(* IEC 61131-3 sources: plc_simulator/plc, 4 files *)

(* ---- types.st ---- *)
USING Siemens.Simatic.Communication.OUC;
USING Siemens.Simatic.Communication.OpenUser;
USING Siemens.Simatic.Communication.MQTT;
USING Siemens.Simatic.Communication.Util;
USING System.Strings;
USING System.Serialization;

/*
#### IO map

1. control box
button: start, stop,reset
led, auto,stop,warn
errormsg

2. belt
motor command: enable, speed
motor state: state, speed

3. sensor
IR
Banner

#### Controller Main Logic
1. running state transition
idle -> running -> suspend -> stop
running -> error -> reset -> running

2. belt layout configuration
graph
link table

2. sequence start

*/

TYPE

    Station_1_Input : STRUCT
        button_1_1_1 : BOOL;
        button_1_1_2 : BOOL;
        button_1_1_3 : BOOL;
        sensor_1_1_1 : BOOL;
        button_1_2_1 : BOOL;
        button_1_2_2 : BOOL;
        button_1_2_3 : BOOL;
        sensor_1_2_1 : DWORD;
        button_1_3_1 : BOOL;
        button_1_3_2 : BOOL;
        button_1_3_3 : BOOL;
        sensor_1_3_1 : DWORD;
        clock : LINT;

    END_STRUCT;
END_TYPE

TYPE
    Station_1_Output : STRUCT
        led_1_1_1 : BOOL;
        led_1_1_2 : BOOL;
        led_1_1_3 : BOOL;
        led_1_2_1 : BOOL;
        led_1_2_2 : BOOL;
        led_1_2_3 : BOOL;
        led_1_3_1 : BOOL;
        led_1_3_2 : BOOL;
        led_1_3_3 : BOOL;

        belt_1_1_1: ARRAY[0..1] of REAL;
        belt_1_1_2: ARRAY[0..1] of REAL;
        belt_1_1_3: ARRAY[0..1] of REAL;
        belt_1_1_4: ARRAY[0..1] of REAL;
        belt_1_1_5: ARRAY[0..1] of REAL;
        // belt_1_1_6: ARRAY[0..1] of REAL;

        belt_1_2_1: ARRAY[0..1] of REAL;
        belt_1_2_2: ARRAY[0..1] of REAL;
        belt_1_2_3: ARRAY[0..1] of REAL;
        belt_1_2_4: ARRAY[0..1] of REAL;
        belt_1_2_5: ARRAY[0..1] of REAL;

        belt_1_3_1: ARRAY[0..1] of REAL;
        belt_1_3_2: ARRAY[0..1] of REAL;
        belt_1_3_3: ARRAY[0..1] of REAL;
        belt_1_3_4: ARRAY[0..1] of REAL;
        belt_1_3_5: ARRAY[0..1] of REAL;

    END_STRUCT;
END_TYPE

(* ---- tcp_client_lib.st ---- *)
USING Siemens.Simatic.Communication.OUC;
USING System;
USING System.Serialization; // For handling byte-to-integer conversions

FUNCTION TcpBlockMove
    VAR_IN_OUT
        source : ARRAY[*] OF BYTE;
        dest : ARRAY[*] OF BYTE;
    END_VAR
    VAR_INPUT
        srcOffset : UDINT;
        dstOffset : UDINT;
        count : UDINT;
    END_VAR
    VAR_TEMP
        I : UDINT;
        srcIdx : DINT;
        dstIdx : DINT;
    END_VAR

    IF count = UDINT#0 THEN
        RETURN;
    END_IF;

    srcIdx := LOWER_BOUND(source, 1) + TO_DINT(srcOffset);
    dstIdx := LOWER_BOUND(dest, 1) + TO_DINT(dstOffset);

    FOR I := UDINT#0 TO count - UDINT#1 DO
        dest[dstIdx] := source[srcIdx];
        srcIdx := srcIdx + DINT#1;
        dstIdx := dstIdx + DINT#1;
    END_FOR;
END_FUNCTION

CLASS TcpClient
    VAR CONSTANT
        MAX_SEND_LENGTH : UINT := UINT#256;
        MAX_RECEIVE_LENGTH : UINT := UINT#256;
    END_VAR

    VAR PUBLIC
        IsConfigured : BOOL := FALSE;
        IsConnected : BOOL := FALSE;

        ConnectDone, ConnectError, ConnectBusy : BOOL;
        ConnectExecute : BOOL;
        ConnectStatus, LastConnectStatus : WORD;
        ConnectAttemptCount, ConnectDoneCount, ConnectErrorCount : UDINT;

        SendDone, SendError, SendBusy : BOOL;
        SendExecute : BOOL;
        SendStatus, LastSendStatus : WORD;
        SendDoneCount, SendErrorCount, DroppedSendCount : UDINT;

        ReceiveNewData, ReceiveError, ReceiveBusy : BOOL;
        ReceiveStatus, LastReceiveStatus : WORD;
        ReceiveLength :INT;
        ReceiveCount, ReceiveErrorCount : UDINT;
        ReceiveBuffer : ARRAY [0..MAX_RECEIVE_LENGTH - UINT#1] OF BYTE;
    END_VAR

    VAR PRIVATE
        config : ConnectionConfiguration;
        connect : Connect;
        send : TcpSend;
        receive : TcpReceive;
        sendTimer : IEC.TON;
        sendPeriod : TIME := T#1S;
        sendBuffer : ARRAY [0..MAX_SEND_LENGTH - UINT#1] OF BYTE;
        sendLength : UDINT := UDINT#0;
        sendQueued : BOOL := FALSE;
        prevConnectExecute : BOOL := FALSE;
           retryTimer : IEC.TON;
    retryDelay : TIME := T#2S;
    forceExecuteLow : BOOL := FALSE;

    END_VAR

    METHOD PUBLIC Configure
        VAR_INPUT
            remoteAddress : Siemens.Simatic.Communication.IPConfiguration.IPv4;
            remotePort : UINT;
            connectionID : WORD := WORD#1;
            hardwareID : UINT := UINT#64;
            period : TIME := T#1S;
        END_VAR

        IF NOT IsConfigured THEN
            config.HardwareID := hardwareID;
            config.ConnectionID := connectionID;
            config.RemoteAddress := remoteAddress;
            config.RemotePort := remotePort;
            sendPeriod := period;
            IsConfigured := TRUE;
        END_IF;
    END_METHOD

    METHOD PUBLIC QueueSend
        VAR_INPUT
            dataLength : UDINT;
        END_VAR
        VAR_IN_OUT
            data : ARRAY[*] OF BYTE;
        END_VAR

        IF (dataLength + UDINT#8) > TO_UDINT(MAX_SEND_LENGTH) THEN
            DroppedSendCount := DroppedSendCount + UDINT#1;
            RETURN;
        END_IF;

        IF SendBusy THEN
            DroppedSendCount := DroppedSendCount + UDINT#1;
            RETURN;
        END_IF;

        sendLength := dataLength + UDINT#8;

        // Fixed magic marker 16#12345678, followed by little-endian UDINT payload length.
        sendBuffer[0] := BYTE#16#12;
        sendBuffer[1] := BYTE#16#34;
        sendBuffer[2] := BYTE#16#56;
        sendBuffer[3] := BYTE#16#78;
        sendBuffer[4] := TO_BYTE(TO_DWORD(dataLength) AND DWORD#16#FF);
        sendBuffer[5] := TO_BYTE(SHR(TO_DWORD(dataLength), USINT#8) AND DWORD#16#FF);
        sendBuffer[6] := TO_BYTE(SHR(TO_DWORD(dataLength), USINT#16) AND DWORD#16#FF);
        sendBuffer[7] := TO_BYTE(SHR(TO_DWORD(dataLength), USINT#24) AND DWORD#16#FF);

        TcpBlockMove(
            source := data,
            dest := sendBuffer,
            srcOffset := UDINT#0,
            dstOffset := UDINT#8,
            count := dataLength
        );

        sendQueued := TRUE;
    END_METHOD

    METHOD PUBLIC Run

        VAR_TEMP
            recv_len : udint;
            END_VAR

// in Run():
IF ConnectError THEN
    forceExecuteLow := TRUE;
    retryTimer(IN := TRUE, PT := retryDelay);
ELSIF retryTimer.Q THEN
    forceExecuteLow := FALSE;
    retryTimer(IN := FALSE);
END_IF;

ConnectExecute := NOT IsConnected AND NOT connect.busy AND NOT forceExecuteLow;

        IF NOT IsConfigured THEN
            RETURN;
        END_IF;

        // ConnectExecute := NOT IsConnected AND NOT connect.busy;
        IF ConnectExecute AND NOT prevConnectExecute THEN
            ConnectAttemptCount := ConnectAttemptCount + UDINT#1;
        END_IF;
        prevConnectExecute := ConnectExecute;

        // connect(
        // execute := NOT IsConnected AND NOT connect.busy,
        // connectionID := config.ConnectionID,
        // connectionConfiguration := config,
        // done => ConnectDone,
        //     busy => ConnectBusy,
        //     error => ConnectError,
        //     status => ConnectStatus
        // );

        connect(
            execute := ConnectExecute,
            connectionID := config.ConnectionID,
            connectionConfiguration := config,
            done => ConnectDone,
            busy => ConnectBusy,
            error => ConnectError,
            status => ConnectStatus
        );

        IF ConnectStatus <> WORD#16#7000 THEN
            LastConnectStatus := ConnectStatus;
        END_IF;

        IF ConnectDone THEN
            ConnectDoneCount := ConnectDoneCount + UDINT#1;
            IsConnected := TRUE;
        END_IF;

        IF ConnectError THEN
            ConnectErrorCount := ConnectErrorCount + UDINT#1;
        END_IF;

        sendTimer(IN := IsConnected AND sendQueued AND NOT sendTimer.Q, PT := sendPeriod);
        SendExecute := IsConnected AND sendQueued AND sendTimer.Q AND NOT send.busy;

        send(
            execute := SendExecute,
            connectionID := config.ConnectionID,
            length := sendLength,
            data := sendBuffer,
            done => SendDone,
            busy => SendBusy,
            error => SendError,
            status => SendStatus
        );

        IF SendStatus <> WORD#16#7000 THEN
            LastSendStatus := SendStatus;
        END_IF;

        IF SendDone THEN
            SendDoneCount := SendDoneCount + UDINT#1;
        END_IF;

        IF SendError THEN
            SendErrorCount := SendErrorCount + UDINT#1;
        END_IF;
        receive(
            enable := IsConnected,
            connectionID := config.ConnectionID,
            adhocMode := TRUE,
            data := ReceiveBuffer,
            length := MAX_RECEIVE_LENGTH,

            newDataReceived => ReceiveNewData,
            receivedLength =>  recv_len,
            busy => ReceiveBusy,
            error => ReceiveError,
            status => ReceiveStatus
        );

        IF ReceiveNewData THEN
            ReceiveLength := TO_INT(recv_len);
        ELSE
            ReceiveLength := INT#0;
        END_IF;

        IF ReceiveStatus <> WORD#16#7000 THEN
            LastReceiveStatus := ReceiveStatus;
        END_IF;

        IF ReceiveNewData THEN
            ReceiveCount := ReceiveCount + UDINT#1;
        END_IF;

        IF ReceiveError THEN
            ReceiveErrorCount := ReceiveErrorCount + UDINT#1;
        END_IF;
    END_METHOD
END_CLASS

CLASS TCP_StreamParser1

    VAR CONSTANT
        BUFFER_LENGTH : INT := 4095;
        PAYLOAD_LENGTH : INT := 2048;

        // Instance of your TRCV or communication interface
        // e.g., MyTrcvInstance : TRCV;
    END_VAR

    VAR
        // Adjust buffer size depending on your largest expected payload + 8 byte header
        Buffer : Array[0..BUFFER_LENGTH] Of Byte;
        BufferLength : Int := 0; // Tracks current number of valid bytes in Buffer

    END_VAR

    VAR PUBLIC
        // Parsing variables
        // i : Int := 0;
        MagicFound : Bool := False;
        MarkerIndex : Int := 0;
        PayloadLength : DInt := 0;
        TotalPacketSize : Int := 0;

        // Output/Export extracted data
        PayloadReady : Bool := False;
        ExtractedPayload : Array[0..PAYLOAD_LENGTH] Of Byte;
        ExtractedLength : Int := 0;
    END_VAR

    METHOD PUBLIC Execute
        VAR
            MoveIndex : Int;

        END_VAR
        VAR_IN_OUT
           // Temp array to capture immediate cycle data from network
            RxTemp : Array[*] Of Byte;
            RxCount : Int;
        END_VAR
        VAR_TEMP
            i : int;

        END_VAR

        PayloadReady := False; // Reset flag every cycle

        // 1. SIMULATED/ACTUAL RECV CALL: Fetch raw data from network interface
        // Replace this block with your actual TRCV logic
        // TRCV_Instance(RCV:=RxTemp, ...NDR=>DataReady, LEN=>RxCount);

        // If data arrived this cycle, append it to our main stream buffer
        IF RxCount > 0 THEN
            // Ensure we don't overflow our main stream buffer
            IF (BufferLength + RxCount) <= 4096 THEN
                // Copy temporary network chunk to the end of our stream buffer
                FOR i := 0 TO RxCount - 1 DO
                    Buffer[BufferLength + i] := RxTemp[i];
                END_FOR;
                BufferLength := BufferLength + RxCount;
            ELSE
                // Handle Buffer Overflow Error here (e.g., reset buffer)
                BufferLength := 0;
            END_IF;
        END_IF;

        // 2. PARSING LOOP: Process buffer continuously until no complete packets remain
        WHILE BufferLength >= 8 DO // Must have at least 8 bytes (4B Magic + 4B Length)

            MagicFound := False;

            // Look for the 4-byte Magic Marker: 0x12345678
            FOR i := 0 TO (BufferLength - 4) DO
                IF Buffer[i] = TO_BYTE(16#12) AND Buffer[i+1] = TO_BYTE(16#34) AND Buffer[i+2] = TO_BYTE(16#56) AND Buffer[i+3] = TO_BYTE(16#78) THEN
                    MagicFound := True;
                    MarkerIndex := i;
                    EXIT; // Found the earliest marker, break FOR loop
                END_IF;
            END_FOR;

            // If magic marker is not anywhere in the buffer, discard junk data safely
            IF NOT MagicFound THEN
                // Keep only the last 3 bytes in case the magic word was split between frames
                IF BufferLength > 3 THEN
                    FOR i := 0 TO 2 DO
                        Buffer[i] := Buffer[BufferLength - 3 + i];
                    END_FOR;
                    BufferLength := 3;
                END_IF;
                EXIT; // Break the WHILE loop, wait for more data
            END_IF;

            // If the magic marker was found deeper in the stream, slide buffer to align to it
            IF MarkerIndex > 0 THEN
                FOR i := 0 TO (BufferLength - 1 - MarkerIndex) DO
                    Buffer[i] := Buffer[MarkerIndex + i];
                END_FOR;
                BufferLength := BufferLength - MarkerIndex;
            END_IF;

            // Double check if we still have the full 8 bytes header after realignment
            IF BufferLength < 8 THEN
                EXIT; // Wait for next cycle data
            END_IF;

            // 3. EXTRACT LENGTH: Deserialize 4 bytes following the magic marker (little-endian)
            // Reconstructs DInt from Buffer[4..7]
            // PayloadLength := TO_DINT(SHL(TO_DWORD(Buffer[4]), UINT#24) OR
            //                  SHL(TO_DWORD(Buffer[5]), UINT#16) OR
            //                  SHL(TO_DWORD(Buffer[6]), UINT#8)  OR
            //                  TO_DWORD(Buffer[7]));

            // Combined safely into a DINT
PayloadLength := TO_DINT(
    TO_DWORD(Buffer[4]) OR
    SHL(TO_DWORD(Buffer[5]), USINT#8) OR
    SHL(TO_DWORD(Buffer[6]), USINT#16) OR
    SHL(TO_DWORD(Buffer[7]), USINT#24)
);

            TotalPacketSize := 8 + TO_INT(PayloadLength);

            // 4. CHECK COMPLETENESS: Ensure the complete payload length has arrived
            IF BufferLength < TotalPacketSize THEN
                EXIT; // Packet incomplete. Stop parsing and wait for the rest of the stream
            END_IF;

            // 5. EXTRACT PAYLOAD: Complete packet found! Copy it to output array
            FOR i := 0 TO TO_INT(PayloadLength) - 1 DO
                ExtractedPayload[i] := Buffer[8 + i];
            END_FOR;

            ExtractedLength := TO_INT(PayloadLength);
            PayloadReady := True; // Signal to consumer logic that data is ready

            // Execute application-specific logic with ExtractedPayload here if needed...

            // 6. SLIDE STREAM BUFFER: Shift remaining trailing data to index 0
            BufferLength := BufferLength - TotalPacketSize;
            IF BufferLength > 0 THEN
                FOR i := 0 TO (BufferLength - 1) DO
                    Buffer[i] := Buffer[TotalPacketSize + i];
                END_FOR;
            END_IF;

        END_WHILE;
    END_METHOD
END_CLASS

CLASS TCP_StreamParser

    VAR CONSTANT
        BUFFER_LENGTH : INT := 4095;
        PAYLOAD_LENGTH : INT := 2048;
        HEADER_SIZE : INT := 8;
    END_VAR

    VAR
        // Persistent internal stream buffer
        Buffer : Array[0..BUFFER_LENGTH] Of Byte;
        BufferLength : Int := 0; // Tracks current number of valid bytes in Buffer
    END_VAR

    VAR PUBLIC
        // Parsing state variables
        MagicFound : Bool := False;
        MarkerIndex : Int := 0;
        PayloadLength : DInt := 0;
        TotalPacketSize : Int := 0;

        // Output / Export data interface
        PayloadReady : Bool := False;
        PayloadReadyCount : Int := 0;

        ExtractedPayload : Array[0..PAYLOAD_LENGTH] Of Byte;
        ExtractedLength : Int := 0;
    END_VAR

    METHOD PUBLIC Execute
        VAR_IN_OUT
            // Dynamic bounds array to safely read variable network chunk sizes
            RxTemp : Array[*] Of Byte;
            RxCount : Int;
        END_VAR

        VAR_TEMP
            i : INT;
            UpperIndexBound : DINT;
        END_VAR

        PayloadReady := False; // Reset flag every cycle

        // 1. APPEND NEW NETWORK DATA TO STREAM BUFFER
        IF RxCount > 0 THEN
            // FIX 1: Dynamically match against the upper bound of the constant size (4095 index = 4096 size)
            IF (BufferLength + RxCount) <= (BUFFER_LENGTH + 1) THEN
                FOR i := 0 TO RxCount - 1 DO
                    Buffer[BufferLength + i] := RxTemp[LOWER_BOUND(RxTemp, 1) + TO_DINT(i)];
                END_FOR;
                BufferLength := BufferLength + RxCount;
            ELSE
                // Buffer Overflow Safety: Wipe pointer to avoid crashing the PLC PLC
                BufferLength := 0;
            END_IF;
        END_IF;

        // 2. PARSING LOOP: Process internal stream buffer
        WHILE BufferLength >= HEADER_SIZE DO

            MagicFound := False;

            // Look for the 4-byte Magic Marker: 0x12345678
            FOR i := 0 TO (BufferLength - 4) DO
                IF Buffer[i] = TO_BYTE(16#12) AND Buffer[i+1] = TO_BYTE(16#34) AND Buffer[i+2] = TO_BYTE(16#56) AND Buffer[i+3] = TO_BYTE(16#78) THEN
                    MagicFound := True;
                    MarkerIndex := i;
                    EXIT; // Found the earliest marker, break FOR loop
                END_IF;
            END_FOR;

            // FIX 2: Handle garbage data or unmatched fragments safely without losing potential split markers
            IF NOT MagicFound THEN
                IF BufferLength > 3 THEN
                    FOR i := 0 TO 2 DO
                        Buffer[i] := Buffer[BufferLength - 3 + i];
                    END_FOR;
                    BufferLength := 3;
                END_IF;
                EXIT; // Force break of WHILE loop to wait for more data
            END_IF;

            // If the magic marker was found deeper in the stream, slide buffer to align to it
            IF MarkerIndex > 0 THEN
                FOR i := 0 TO (BufferLength - 1 - MarkerIndex) DO
                    Buffer[i] := Buffer[MarkerIndex + i];
                END_FOR;
                BufferLength := BufferLength - MarkerIndex;
            END_IF;

            // Re-verify we still have a header window left after shifting
            IF BufferLength < HEADER_SIZE THEN
                EXIT;
            END_IF;

            // 3. EXTRACT LENGTH (little-endian UDINT from fixed magic frame)
            PayloadLength := TO_DINT(
                TO_DWORD(Buffer[4]) OR
                SHL(TO_DWORD(Buffer[5]), USINT#8) OR
                SHL(TO_DWORD(Buffer[6]), USINT#16) OR
                SHL(TO_DWORD(Buffer[7]), USINT#24)
            );

            TotalPacketSize := HEADER_SIZE + TO_INT(PayloadLength);

            // FIX 3: Safety verification against internal memory sizing bounds
            IF TotalPacketSize > (BUFFER_LENGTH + 1) OR TO_INT(PayloadLength) > (PAYLOAD_LENGTH + 1) THEN
                // Protocol violation or data corruption occurred. Flush buffer to reset syncing alignment.
                BufferLength := 0;
                EXIT;
            END_IF;

            // 4. CHECK COMPLETENESS: Ensure full payload has arrived
            IF BufferLength < TotalPacketSize THEN
                EXIT; // Stop parsing this cycle, await more TCP fragments
            END_IF;

            // 5. EXTRACT PAYLOAD
            FOR i := 0 TO TO_INT(PayloadLength) - 1 DO
                ExtractedPayload[i] := Buffer[HEADER_SIZE + i];
            END_FOR;

            ExtractedLength := TO_INT(PayloadLength);
            PayloadReady := True;

            IF PayloadReady THEN
                PayloadReadyCount := PayloadReadyCount + 1;
            END_IF;

            // FIX 4: Put application callback trigger HERE if handling multiple frames in 1 cycle
            // This ensures every parsed message gets intercepted before being overwritten below

            // 6. SLIDE STREAM BUFFER AHEAD
            BufferLength := BufferLength - TotalPacketSize;
            IF BufferLength > 0 THEN
                FOR i := 0 TO (BufferLength - 1) DO
                    Buffer[i] := Buffer[TotalPacketSize + i];
                END_FOR;
            END_IF;

            // FIX 5: Prevent infinite loops if a corrupted packet sets PayloadLength to 0
            IF TotalPacketSize <= HEADER_SIZE THEN
                BufferLength := 0;
                EXIT;
            END_IF;

        END_WHILE;
    END_METHOD
END_CLASS

(* ---- types-generated.st ---- *)
// -----------------------------------------------------------------------------
// <auto-generated>
// Generated by tools/generate_st_serde.py. Do not edit by hand.
// -----------------------------------------------------------------------------
USING System.Serialization;
USING System.BitAccess;

// Generated from src/types.st:15
// Byte mapping, relative to startOffset:
//   button_1_1_1 -> byte 0, bit 0
//   button_1_1_2 -> byte 0, bit 1
//   button_1_1_3 -> byte 0, bit 2
//   sensor_1_1_1 -> byte 0, bit 3
//   button_1_2_1 -> byte 0, bit 4
//   button_1_2_2 -> byte 0, bit 5
//   button_1_2_3 -> byte 0, bit 6
//   <padding> -> byte 0, bits 7..7
//   sensor_1_2_1 -> bytes 1..4
//   button_1_3_1 -> byte 5, bit 0
//   button_1_3_2 -> byte 5, bit 1
//   button_1_3_3 -> byte 5, bit 2
//   <padding> -> byte 5, bits 3..7
//   sensor_1_3_1 -> bytes 6..9
//   clock -> bytes 10..17
// Total serialized size: 18 byte(s)
FUNCTION DeserializeFromBytes : UDINT
    VAR_INPUT
        startOffset : UDINT := UDINT#0;
    END_VAR
    VAR_IN_OUT
        source : ARRAY[*] OF BYTE;
        value : Station_1_Input;
    END_VAR
    VAR_TEMP
        offset : UDINT;
        baseIdx : DINT;
        byteIdx : DINT;
    END_VAR

    offset := startOffset;
    baseIdx := LOWER_BOUND(source, 1);
    byteIdx := baseIdx + TO_DINT(offset);
    value.button_1_1_1 := GetBit(source[byteIdx], USINT#0);
    value.button_1_1_2 := GetBit(source[byteIdx], USINT#1);
    value.button_1_1_3 := GetBit(source[byteIdx], USINT#2);
    value.sensor_1_1_1 := GetBit(source[byteIdx], USINT#3);
    value.button_1_2_1 := GetBit(source[byteIdx], USINT#4);
    value.button_1_2_2 := GetBit(source[byteIdx], USINT#5);
    value.button_1_2_3 := GetBit(source[byteIdx], USINT#6);
    offset := offset + UDINT#1;
    offset := Deserialize(offset, source, value.sensor_1_2_1);
    byteIdx := baseIdx + TO_DINT(offset);
    value.button_1_3_1 := GetBit(source[byteIdx], USINT#0);
    value.button_1_3_2 := GetBit(source[byteIdx], USINT#1);
    value.button_1_3_3 := GetBit(source[byteIdx], USINT#2);
    offset := offset + UDINT#1;
    offset := Deserialize(offset, source, value.sensor_1_3_1);
    offset := Deserialize(offset, source, value.clock);
    DeserializeFromBytes := offset;
END_FUNCTION

FUNCTION SerializeToBytes : UDINT
    VAR_INPUT
        startOffset : UDINT := UDINT#0;
    END_VAR
    VAR_IN_OUT
        value : Station_1_Input;
        dest : ARRAY[*] OF BYTE;
    END_VAR
    VAR_TEMP
        offset : UDINT;
        baseIdx : DINT;
        byteIdx : DINT;
    END_VAR

    offset := startOffset;
    baseIdx := LOWER_BOUND(dest, 1);
    byteIdx := baseIdx + TO_DINT(offset);
    dest[byteIdx] := BYTE#16#00;
    dest[byteIdx] := SetBit(value := dest[byteIdx], index := USINT#0, bitValue := value.button_1_1_1);
    dest[byteIdx] := SetBit(value := dest[byteIdx], index := USINT#1, bitValue := value.button_1_1_2);
    dest[byteIdx] := SetBit(value := dest[byteIdx], index := USINT#2, bitValue := value.button_1_1_3);
    dest[byteIdx] := SetBit(value := dest[byteIdx], index := USINT#3, bitValue := value.sensor_1_1_1);
    dest[byteIdx] := SetBit(value := dest[byteIdx], index := USINT#4, bitValue := value.button_1_2_1);
    dest[byteIdx] := SetBit(value := dest[byteIdx], index := USINT#5, bitValue := value.button_1_2_2);
    dest[byteIdx] := SetBit(value := dest[byteIdx], index := USINT#6, bitValue := value.button_1_2_3);
    offset := offset + UDINT#1;
    offset := Serialize(offset, value.sensor_1_2_1, dest);
    byteIdx := baseIdx + TO_DINT(offset);
    dest[byteIdx] := BYTE#16#00;
    dest[byteIdx] := SetBit(value := dest[byteIdx], index := USINT#0, bitValue := value.button_1_3_1);
    dest[byteIdx] := SetBit(value := dest[byteIdx], index := USINT#1, bitValue := value.button_1_3_2);
    dest[byteIdx] := SetBit(value := dest[byteIdx], index := USINT#2, bitValue := value.button_1_3_3);
    offset := offset + UDINT#1;
    offset := Serialize(offset, value.sensor_1_3_1, dest);
    offset := Serialize(offset, value.clock, dest);
    SerializeToBytes := offset;
END_FUNCTION

// Generated from src/types.st:35
// Byte mapping, relative to startOffset:
//   led_1_1_1 -> byte 0, bit 0
//   led_1_1_2 -> byte 0, bit 1
//   led_1_1_3 -> byte 0, bit 2
//   led_1_2_1 -> byte 0, bit 3
//   led_1_2_2 -> byte 0, bit 4
//   led_1_2_3 -> byte 0, bit 5
//   led_1_3_1 -> byte 0, bit 6
//   led_1_3_2 -> byte 0, bit 7
//   led_1_3_3 -> byte 1, bit 0
//   <padding> -> byte 1, bits 1..7
//   belt_1_1_1[0] -> bytes 2..5
//   belt_1_1_1[1] -> bytes 6..9
//   belt_1_1_2[0] -> bytes 10..13
//   belt_1_1_2[1] -> bytes 14..17
//   belt_1_1_3[0] -> bytes 18..21
//   belt_1_1_3[1] -> bytes 22..25
//   belt_1_1_4[0] -> bytes 26..29
//   belt_1_1_4[1] -> bytes 30..33
//   belt_1_1_5[0] -> bytes 34..37
//   belt_1_1_5[1] -> bytes 38..41
//   belt_1_2_1[0] -> bytes 42..45
//   belt_1_2_1[1] -> bytes 46..49
//   belt_1_2_2[0] -> bytes 50..53
//   belt_1_2_2[1] -> bytes 54..57
//   belt_1_2_3[0] -> bytes 58..61
//   belt_1_2_3[1] -> bytes 62..65
//   belt_1_2_4[0] -> bytes 66..69
//   belt_1_2_4[1] -> bytes 70..73
//   belt_1_2_5[0] -> bytes 74..77
//   belt_1_2_5[1] -> bytes 78..81
//   belt_1_3_1[0] -> bytes 82..85
//   belt_1_3_1[1] -> bytes 86..89
//   belt_1_3_2[0] -> bytes 90..93
//   belt_1_3_2[1] -> bytes 94..97
//   belt_1_3_3[0] -> bytes 98..101
//   belt_1_3_3[1] -> bytes 102..105
//   belt_1_3_4[0] -> bytes 106..109
//   belt_1_3_4[1] -> bytes 110..113
//   belt_1_3_5[0] -> bytes 114..117
//   belt_1_3_5[1] -> bytes 118..121
// Total serialized size: 122 byte(s)
FUNCTION DeserializeFromBytes : UDINT
    VAR_INPUT
        startOffset : UDINT := UDINT#0;
    END_VAR
    VAR_IN_OUT
        source : ARRAY[*] OF BYTE;
        value : Station_1_Output;
    END_VAR
    VAR_TEMP
        offset : UDINT;
        baseIdx : DINT;
        byteIdx : DINT;
    END_VAR

    offset := startOffset;
    baseIdx := LOWER_BOUND(source, 1);
    byteIdx := baseIdx + TO_DINT(offset);
    value.led_1_1_1 := GetBit(source[byteIdx], USINT#0);
    value.led_1_1_2 := GetBit(source[byteIdx], USINT#1);
    value.led_1_1_3 := GetBit(source[byteIdx], USINT#2);
    value.led_1_2_1 := GetBit(source[byteIdx], USINT#3);
    value.led_1_2_2 := GetBit(source[byteIdx], USINT#4);
    value.led_1_2_3 := GetBit(source[byteIdx], USINT#5);
    value.led_1_3_1 := GetBit(source[byteIdx], USINT#6);
    value.led_1_3_2 := GetBit(source[byteIdx], USINT#7);
    offset := offset + UDINT#1;
    byteIdx := baseIdx + TO_DINT(offset);
    value.led_1_3_3 := GetBit(source[byteIdx], USINT#0);
    offset := offset + UDINT#1;
    offset := Deserialize(offset, source, value.belt_1_1_1[0]);
    offset := Deserialize(offset, source, value.belt_1_1_1[1]);
    offset := Deserialize(offset, source, value.belt_1_1_2[0]);
    offset := Deserialize(offset, source, value.belt_1_1_2[1]);
    offset := Deserialize(offset, source, value.belt_1_1_3[0]);
    offset := Deserialize(offset, source, value.belt_1_1_3[1]);
    offset := Deserialize(offset, source, value.belt_1_1_4[0]);
    offset := Deserialize(offset, source, value.belt_1_1_4[1]);
    offset := Deserialize(offset, source, value.belt_1_1_5[0]);
    offset := Deserialize(offset, source, value.belt_1_1_5[1]);
    offset := Deserialize(offset, source, value.belt_1_2_1[0]);
    offset := Deserialize(offset, source, value.belt_1_2_1[1]);
    offset := Deserialize(offset, source, value.belt_1_2_2[0]);
    offset := Deserialize(offset, source, value.belt_1_2_2[1]);
    offset := Deserialize(offset, source, value.belt_1_2_3[0]);
    offset := Deserialize(offset, source, value.belt_1_2_3[1]);
    offset := Deserialize(offset, source, value.belt_1_2_4[0]);
    offset := Deserialize(offset, source, value.belt_1_2_4[1]);
    offset := Deserialize(offset, source, value.belt_1_2_5[0]);
    offset := Deserialize(offset, source, value.belt_1_2_5[1]);
    offset := Deserialize(offset, source, value.belt_1_3_1[0]);
    offset := Deserialize(offset, source, value.belt_1_3_1[1]);
    offset := Deserialize(offset, source, value.belt_1_3_2[0]);
    offset := Deserialize(offset, source, value.belt_1_3_2[1]);
    offset := Deserialize(offset, source, value.belt_1_3_3[0]);
    offset := Deserialize(offset, source, value.belt_1_3_3[1]);
    offset := Deserialize(offset, source, value.belt_1_3_4[0]);
    offset := Deserialize(offset, source, value.belt_1_3_4[1]);
    offset := Deserialize(offset, source, value.belt_1_3_5[0]);
    offset := Deserialize(offset, source, value.belt_1_3_5[1]);
    DeserializeFromBytes := offset;
END_FUNCTION

FUNCTION SerializeToBytes : UDINT
    VAR_INPUT
        startOffset : UDINT := UDINT#0;
    END_VAR
    VAR_IN_OUT
        value : Station_1_Output;
        dest : ARRAY[*] OF BYTE;
    END_VAR
    VAR_TEMP
        offset : UDINT;
        baseIdx : DINT;
        byteIdx : DINT;
    END_VAR

    offset := startOffset;
    baseIdx := LOWER_BOUND(dest, 1);
    byteIdx := baseIdx + TO_DINT(offset);
    dest[byteIdx] := BYTE#16#00;
    dest[byteIdx] := SetBit(value := dest[byteIdx], index := USINT#0, bitValue := value.led_1_1_1);
    dest[byteIdx] := SetBit(value := dest[byteIdx], index := USINT#1, bitValue := value.led_1_1_2);
    dest[byteIdx] := SetBit(value := dest[byteIdx], index := USINT#2, bitValue := value.led_1_1_3);
    dest[byteIdx] := SetBit(value := dest[byteIdx], index := USINT#3, bitValue := value.led_1_2_1);
    dest[byteIdx] := SetBit(value := dest[byteIdx], index := USINT#4, bitValue := value.led_1_2_2);
    dest[byteIdx] := SetBit(value := dest[byteIdx], index := USINT#5, bitValue := value.led_1_2_3);
    dest[byteIdx] := SetBit(value := dest[byteIdx], index := USINT#6, bitValue := value.led_1_3_1);
    dest[byteIdx] := SetBit(value := dest[byteIdx], index := USINT#7, bitValue := value.led_1_3_2);
    offset := offset + UDINT#1;
    byteIdx := baseIdx + TO_DINT(offset);
    dest[byteIdx] := BYTE#16#00;
    dest[byteIdx] := SetBit(value := dest[byteIdx], index := USINT#0, bitValue := value.led_1_3_3);
    offset := offset + UDINT#1;
    offset := Serialize(offset, value.belt_1_1_1[0], dest);
    offset := Serialize(offset, value.belt_1_1_1[1], dest);
    offset := Serialize(offset, value.belt_1_1_2[0], dest);
    offset := Serialize(offset, value.belt_1_1_2[1], dest);
    offset := Serialize(offset, value.belt_1_1_3[0], dest);
    offset := Serialize(offset, value.belt_1_1_3[1], dest);
    offset := Serialize(offset, value.belt_1_1_4[0], dest);
    offset := Serialize(offset, value.belt_1_1_4[1], dest);
    offset := Serialize(offset, value.belt_1_1_5[0], dest);
    offset := Serialize(offset, value.belt_1_1_5[1], dest);
    offset := Serialize(offset, value.belt_1_2_1[0], dest);
    offset := Serialize(offset, value.belt_1_2_1[1], dest);
    offset := Serialize(offset, value.belt_1_2_2[0], dest);
    offset := Serialize(offset, value.belt_1_2_2[1], dest);
    offset := Serialize(offset, value.belt_1_2_3[0], dest);
    offset := Serialize(offset, value.belt_1_2_3[1], dest);
    offset := Serialize(offset, value.belt_1_2_4[0], dest);
    offset := Serialize(offset, value.belt_1_2_4[1], dest);
    offset := Serialize(offset, value.belt_1_2_5[0], dest);
    offset := Serialize(offset, value.belt_1_2_5[1], dest);
    offset := Serialize(offset, value.belt_1_3_1[0], dest);
    offset := Serialize(offset, value.belt_1_3_1[1], dest);
    offset := Serialize(offset, value.belt_1_3_2[0], dest);
    offset := Serialize(offset, value.belt_1_3_2[1], dest);
    offset := Serialize(offset, value.belt_1_3_3[0], dest);
    offset := Serialize(offset, value.belt_1_3_3[1], dest);
    offset := Serialize(offset, value.belt_1_3_4[0], dest);
    offset := Serialize(offset, value.belt_1_3_4[1], dest);
    offset := Serialize(offset, value.belt_1_3_5[0], dest);
    offset := Serialize(offset, value.belt_1_3_5[1], dest);
    SerializeToBytes := offset;
END_FUNCTION

(* ---- tcp_client.st ---- *)
USING Siemens.Simatic.Communication.OUC;

USING Siemens.Simatic.Communication.OpenUser;
USING Siemens.Simatic.Communication.MQTT;
USING Siemens.Simatic.Communication.Util;
USING System.Strings;
USING System.Serialization;

USING Simatic.Ax.IO.Input;
USING Simatic.Ax.IO.Output;

CONFIGURATION myPLC
    TASK Main(Interval := T#10ms, Priority := 16);
    PROGRAM P2 WITH Main : CommunicationProgram;

    VAR_GLOBAL
        sDONE, sERROR : BOOL;
        sSTATUS : WORD;
        sSendDONE, sSendERROR : BOOL;
        sSendSTATUS : WORD;
        sSendExecute, sSendBusy : BOOL;
        sSendDoneCount, sSendErrorCount : UDINT;
        sLastSendSTATUS : WORD;
        sReceiveNewData, sReceiveBusy, sReceiveERROR : BOOL;
        sReceiveSTATUS, sLastReceiveSTATUS : WORD;
        sReceiveLength : INT;
        sReceiveCount, sReceiveErrorCount : UDINT;
        sReceiveBuffer : ARRAY [0..63] OF BYTE;
        sCycleCount : UDINT;
        sConnectAttemptCount, sConnectDoneCount, sConnectErrorCount : UDINT;
        sLastConnectSTATUS : WORD;
        sConnectExecute, sConnectBusy : BOOL;
        sConnected : BOOL;
                tcpClient : TcpClient;
        tcp_praser:TCP_StreamParser;

    END_VAR
END_CONFIGURATION

PROGRAM CommunicationProgram
    VAR_EXTERNAL
        sDONE, sERROR : BOOL;
        sSTATUS : WORD;
        sSendDONE, sSendERROR : BOOL;
        sSendSTATUS : WORD;
        sSendExecute, sSendBusy : BOOL;
        sSendDoneCount, sSendErrorCount : UDINT;
        sLastSendSTATUS : WORD;
        sReceiveNewData, sReceiveBusy, sReceiveERROR : BOOL;
        sReceiveSTATUS, sLastReceiveSTATUS : WORD;
        sReceiveLength : INT;
        sReceiveCount, sReceiveErrorCount : UDINT;
        sReceiveBuffer : ARRAY [0..63] OF BYTE;
        sCycleCount : UDINT;
        sConnectAttemptCount, sConnectDoneCount, sConnectErrorCount : UDINT;
        sLastConnectSTATUS : WORD;
        sConnectExecute, sConnectBusy : BOOL;
        sConnected : BOOL;

        MI_staion_1: Station_1_Input;
        MO_staion_1: Station_1_Output;
       MO_pubBuffer: ARRAY[0..UDINT#255] OF BYTE;
       MO_pubMirror: Station_1_Output;

       MO_pubLen: UDINT;

    END_VAR

    VAR_EXTERNAL
                tcpClient : TcpClient;
        tcp_praser:TCP_StreamParser;
        END_VAR
    VAR
        // tcpClient : TcpClient;
        // tcp_praser:TCP_StreamParser;
        brokerIp : Siemens.Simatic.Communication.IPConfiguration.IPv4 := [BYTE#192, BYTE#168, BYTE#10, BYTE#11];
        data : ARRAY [0..4] OF BYTE := [BYTE#72, BYTE#69, BYTE#76, BYTE#76, BYTE#79];
        payloadQueued : BOOL := FALSE;
    END_VAR
    VAR_TEMP
        i : DINT;
    END_VAR

    sCycleCount := sCycleCount + UDINT#1;

    tcpClient.Configure(
        remoteAddress := brokerIp,
        remotePort := UINT#5001,
        connectionID := WORD#2,
        hardwareID := UINT#64,
        period := T#10MS
    );

    // IF NOT payloadQueued THEN
    //     tcpClient.QueueSend(
    //         data := data,
    //         dataLength := UDINT#5
    //     );
    //     payloadQueued := TRUE;
    // END_IF;

    tcpClient.Run();

    sDONE := tcpClient.ConnectDone;
    sERROR := tcpClient.ConnectError;
    sSTATUS := tcpClient.ConnectStatus;
    sConnectExecute := tcpClient.ConnectExecute;
    sConnectBusy := tcpClient.ConnectBusy;
    sConnectAttemptCount := tcpClient.ConnectAttemptCount;
    sConnectDoneCount := tcpClient.ConnectDoneCount;
    sConnectErrorCount := tcpClient.ConnectErrorCount;
    sLastConnectSTATUS := tcpClient.LastConnectStatus;
    sConnected := tcpClient.IsConnected;

    sSendDONE := tcpClient.SendDone;
    sSendERROR := tcpClient.SendError;
    sSendSTATUS := tcpClient.SendStatus;
    sSendExecute := tcpClient.SendExecute;
    sSendBusy := tcpClient.SendBusy;
    sSendDoneCount := tcpClient.SendDoneCount;
    sSendErrorCount := tcpClient.SendErrorCount;
    sLastSendSTATUS := tcpClient.LastSendStatus;

    sReceiveNewData := tcpClient.ReceiveNewData;
    sReceiveBusy := tcpClient.ReceiveBusy;
    sReceiveERROR := tcpClient.ReceiveError;
    sReceiveSTATUS := tcpClient.ReceiveStatus;
    sLastReceiveSTATUS := tcpClient.LastReceiveStatus;
    sReceiveLength := tcpClient.ReceiveLength;
    sReceiveCount := tcpClient.ReceiveCount;
    sReceiveErrorCount := tcpClient.ReceiveErrorCount;

    // FOR i := DINT#0 TO DINT#63 DO
    //     sReceiveBuffer[i] := tcpClient.ReceiveBuffer[i];
    // END_FOR;

    tcp_praser.Execute(tcpClient.ReceiveBuffer, tcpClient.ReceiveLength);

// tcp_praser.ExtractedPayload[0] :=1;

    // DeserializeFromBytes(startOffset := UDINT#0, source := tcpClient.ReceiveBuffer, value := MI_staion_1);

    if tcp_praser.PayloadReady THEN

        DeserializeFromBytes(startOffset := UDINT#0, source := tcp_praser.ExtractedPayload, value := MI_staion_1);
    END_IF;

        if MI_staion_1.button_1_1_1 = TRUE THEN

        MO_staion_1.led_1_1_1 := TRUE;
        MO_staion_1.led_1_1_2 := FALSE;

    MO_staion_1.belt_1_1_1[0] := REAL#1.0;
    MO_staion_1.belt_1_1_2[0] := REAL#1.0;
    MO_staion_1.belt_1_1_3[0] := REAL#1.0;
    MO_staion_1.belt_1_1_4[0] := REAL#1.0;
    MO_staion_1.belt_1_1_5[0] := REAL#1.0;
    else
         MO_staion_1.led_1_1_1 := FALSE;
        MO_staion_1.led_1_1_2 := TRUE;
    MO_staion_1.belt_1_1_1[0] := REAL#0.0;
    MO_staion_1.belt_1_1_2[0] := REAL#0.0;
    MO_staion_1.belt_1_1_3[0] := REAL#0.0;
    MO_staion_1.belt_1_1_4[0] := REAL#0.0;
    MO_staion_1.belt_1_1_5[0] := REAL#0.0;
    END_IF;

    MO_pubLen := SerializeToBytes(
        startOffset := UDINT#0,
        value := MO_staion_1,
        dest := MO_pubBuffer
    );
    DeserializeFromBytes(startOffset := UDINT#0, source := MO_pubBuffer, value := MO_pubMirror);

    tcpClient.QueueSend(
                dataLength := MO_pubLen,
                data := MO_pubBuffer
    );

END_PROGRAM
